// Frozen copy of IAG50cm develop 744020b (before IAG50cm#17), the oracle of IagLibraryMatchesLegacy_Tests. Only the names
// and the two types that moved to BROTLib are changed. Do not change it.
FUNCTION_BLOCK FB_PointingModelInversion744
VAR_INPUT
	HourAngle		: LREAL;
	Declination		: LREAL;
	Altitude		: LREAL;
	Latitude		: LREAL;
	epsilon			: LREAL := 0.25; //iteration accuracy in arcsec
	eRefractionMode	: BROTLib.E_RefractionMode := BROTLib.E_RefractionMode.OLD;	// coefficient set of the forward model (IAG50cm#7)
END_VAR
VAR_OUTPUT
	HourAngle_correction	: LREAL;
	Declination_correction	: LREAL;
	bValid					: BOOL;	// FALSE if the iteration did not converge within epsilon (e.g. altitude too close to the horizon, where the model is chaotic -- see testing/check_pointing_inversion.py). HourAngle_correction/Declination_correction are 0.0 when FALSE.
END_VAR
VAR
	fbpointing : FB_PointingModelForward744;
	d_ha		: LREAL := 0.0;
	d_dec		: LREAL := 0.0;
	d_ha_new	: LREAL := 0.0;
	d_dec_new	: LREAL := 0.0;
	i			: INT;
	
END_VAR

// iterate untill diff < epsilon or i_max=7 is reached
// 5 passes converge to <0.25" for the normal operating envelope (alt >= 3deg);
// see testing/check_pointing_inversion.py. Kept a small margin over the bare minimum.
bValid := FALSE;
FOR i:=0 TO 7 BY 1 DO
	d_ha := d_ha_new;
	d_dec := d_dec_new;
	fbpointing(
		HourAngle := LMOD(HourAngle-d_ha,360),
		Declination:= Declination-d_dec,
		Latitude:= Latitude,
		eRefractionMode := eRefractionMode,
		HourAngle_correction => d_ha_new,
		Declination_correction => d_dec_new
	);
	IF NOT fbpointing.bValid THEN
		EXIT;	// below 1 deg altitude the forward model gives 0 (#134), that is not a converged result
	END_IF
	IF ABS(d_ha - d_ha_new) <= epsilon/3600.0 AND ABS(d_dec - d_dec_new) <= epsilon/3600.0 THEN
		bValid := TRUE;
		EXIT;
	END_IF
END_FOR;
// below alt~2-3deg the map is chaotic and never settles within epsilon (see script above);
// do not hand back whatever the last unconverged pass produced
IF bValid THEN
	HourAngle_correction := d_ha_new;
	Declination_correction := d_dec_new;
ELSE
	HourAngle_correction := 0.0;
	Declination_correction := 0.0;
END_IF

END_FUNCTION_BLOCK

(* stored: Version 1.1.0.1, ProductVersion 3.1.4024.15
   POU FB_PointingModelInversion744: Id {6c0bf817-169f-465b-8447-88c59d8d1690}, SpecialFunc None *)
